Fanuc KAREL source: kt00405.KL

-- PROVISIONAL review KL for V770-1; original PC SHA256 b49ae9d83a2dc34eff216ffbb6b8cec8740836628449fd7e7b34bf9f2ff325b2
-- Incomplete behavior may be omitted. Consult companion uncertainty JSON. Do not deploy.
PROGRAM KT00405
%NOLOCKGROUP
VAR
  R1 : REAL
  I2 : INTEGER
  OUT : BOOLEAN
BEGIN
  -- UNRESOLVED_PC offsets 5-16; opcodes 2E,23
  -- UNRESOLVED_PC offsets 21-32; opcodes 2E,23
  -- UNRESOLVED_PC offsets 37-57; opcodes 21,21,64,71,23
  -- UNRESOLVED_PC offsets 62-66; opcodes 7F
END KT00405
